Staubli VAL3: main.pgx

public program main()
  local bool l_bExit
  local string l_sTColor
  local string l_sEColor
  local num l_nClock
  local string l_sFColor
  local string l_sLstMsg
begin
  do
    if util:sPage!="message"
      util:sPage="message"
      call util:loadingPage()
      call bind()
      userPage(util:sPage)
      nMsgType=0
      call initMsg()
      call rs:getLog(sRobotMsg,nMsgType)
      userPageSet("message","btnAllMsg","style.backgroundColor","#33FF33")
      userPageSet("message","btnRobotMsg","style.backgroundColor","#FFFFFF")
      userPageSet("message","btnTrajMsg","style.backgroundColor","#FFFFFF")
      sCurrentMsg=""
    endIf
    if sCurrentMsg!=l_sLstMsg
      l_sLstMsg=sCurrentMsg
      popUpMsg(l_sLstMsg)
      sCurrentMsg=l_sLstMsg=""
    endIf
    if bBack
      bBack=false
      l_bExit=true
    endIf
    delay(0.2)
  until l_bExit==true
end
